Staubli VAL3: stop.pgx

program stop()
begin
  //kill all task
  taskKill("Reset")
  taskKill("Start")
  taskKill("Stop")
  taskKill("cycleCtrl")
  taskKill("Zones")
  taskKill("Main")
  taskKill("StatusRobot")
  //
  stopMove()
  resetMotion()
  disablePower()
end
